Staubli VAL3: hmiConfirm.pgx

public program hmiConfirm(string x_sMsg, string x_sMsgType, bool& x_bOK)
  local string l_sMsg
  local bool l_bOut
begin
  switch sLanguage
    case "english"
      l_sMsg=sAlertEN[x_sMsg]
    break
    case "chinese"
      l_sMsg=sAlertCN[x_sMsg]
    break
  endSwitch
  //*************************************************************
  utCtn_Message.Common.sSource="Page_Container_Confirm.html"
  utTxt_popUpMsg.Common.sValue=l_sMsg
  //*************************************************************
  switch x_sMsgType
    case "info"
      utTxt_popUpMsg.Appearance.sBackgroundColour="#7C95FF"
    break
    //
    case "warning"
      utTxt_popUpMsg.Appearance.sBackgroundColour="#EEFB45"
    break
    //
    case "confirm"
      utTxt_popUpMsg.Appearance.sBackgroundColour="#FFFFFF"
    break
    //
    default
      utTxt_popUpMsg.Appearance.sBackgroundColour="#ADADB2"
    break
  endSwitch
  delay(0.2)
  //
  utCtn_Message.Appearance.bVisibility=true
  //
  utBtn_Yes.Events.bClick=false
  utBtn_No.Events.bClick=false
  l_bOut=false
  do
    if utBtn_Yes.Events.bClick==true
      utBtn_Yes.Events.bClick=false
      l_bOut=true
      x_bOK=true
    elseIf utBtn_No.Events.bClick==true
      utBtn_No.Events.bClick=false
      l_bOut=true
      x_bOK=false
    endIf
  until l_bOut
  delay(0)
  utCtn_Message.Appearance.bVisibility=false
end
